(*
SPDX-FileCopyrightText: © 2026 Oleksandr Tiutyk <trofimich@gmail.com>
SPDX-License-Identifier: MIT
License: https://opensource.org/license/mit
*)

(*!
<summary>Writes run summaries and leaf failures to the ADS log.</summary>
<description>
Use in one task without reentry. The ADS backend has no established concurrent-call guarantee, even for
separate reporter instances. For multiple tasks use per-task in-memory reports or a synchronized backend.
Each callback submits at most one record. The ADS completion record includes counts and the first failed leaf name.
LastRunSummary includes the first failed leaf name and a bounded
version of its diagnostic. The summary and failed log writes are observable after the run. A failed
write does not change the test outcome. Individual ADS failure records are capped at 200 wide characters.
ReportRunStart clears all observations before attempting the start message.
</description>
*)

{attribute 'no_explicit_call' := 'do not call this function block directly'}
FUNCTION_BLOCK AdsLogReporter EXTENDS TOF_Core.Object IMPLEMENTS ITestReporter
VAR_STAT
	_ClassName : STRING := __POUNAME();
END_VAR
VAR
	_AdsLogger : TOF_Core.AdsLogger;
	_FirstFailureName : WSTRING;
	_FirstFailureDiagnostic : WSTRING(255);
	_LastRunSummary : TOF_Core.ERROR_MESSAGE;
	_FailedLogWriteCount : UDINT;
	_LastLogFailureMessage : TOF_Core.ERROR_MESSAGE;
END_VAR

(*!
<summary>Provides the implementation class name.</summary>
*)
{attribute 'monitoring' := 'call'}
PROPERTY ClassName : REFERENCE TO STRING
GET
ClassName REF= _ClassName;
END_GET
END_PROPERTY

(*!
<summary>Counts start, result and summary writes for which TryLogMessage returned FALSE.</summary>
<description>The count resets at ReportRunStart. A successful write does not confirm display in XAE.</description>
*)
{attribute 'monitoring' := 'call'}
PROPERTY FailedLogWriteCount : UDINT
GET
FailedLogWriteCount := _FailedLogWriteCount;
END_GET
END_PROPERTY

(*!
<summary>Borrows the last message whose ADS logger call returned FALSE.</summary>
<description>Empty until a write fails in the current run. Callers must not modify the returned storage.</description>
*)
{attribute 'monitoring' := 'call'}
PROPERTY LastLogFailureMessage : REFERENCE TO TOF_Core.ERROR_MESSAGE
GET
LastLogFailureMessage REF= _LastLogFailureMessage;
END_GET
END_PROPERTY

(*!
<summary>Borrows the summary created at ReportRunEnd regardless of its ADS write status.</summary>
<description>Empty after ReportRunStart until ReportRunEnd. Callers must not modify the returned storage.</description>
*)
{attribute 'monitoring' := 'call'}
PROPERTY LastRunSummary : REFERENCE TO TOF_Core.ERROR_MESSAGE
GET
LastRunSummary REF= _LastRunSummary;
END_GET
END_PROPERTY

(*!
<summary>Submits one ADS message and records a FALSE result from the logger.</summary>
<description>The count saturates at the largest UDINT. The copied text remains available until the next start.</description>
*)
METHOD PRIVATE logMessage
VAR_INPUT
	category : TOF_Core.LOG_CATEGORY;
END_VAR
VAR_IN_OUT CONSTANT
	message : TOF_Core.ERROR_MESSAGE;
END_VAR
IF TryWriteMessage(category := category, message := message) THEN
	RETURN;
END_IF

IF _FailedLogWriteCount < TOF_Core.UnsignedInt32.MAX_VALUE THEN
	_FailedLogWriteCount := _FailedLogWriteCount + 1;
END_IF

_LastLogFailureMessage := message;
END_METHOD

(*!
<summary>Provides the library namespace.</summary>
*)
{attribute 'monitoring' := 'call'}
PROPERTY NamespaceName : REFERENCE TO STRING
GET
NamespaceName REF= CurrentNamespace.Name;
END_GET
END_PROPERTY

(*!
<summary>Logs leaf counts and the first failed leaf name and retains its diagnostic for online inspection.</summary>
<description>The retained summary also includes a bounded first-failure diagnostic and survives a rejected ADS write.</description>
*)
METHOD ReportRunEnd
VAR_INPUT
	totalTests : TOF_Core.DINT_LENGTH;
	passedTests : TOF_Core.DINT_LENGTH;
	failedTests : TOF_Core.DINT_LENGTH;
	skippedTests : TOF_Core.DINT_LENGTH;
	duration : TIME;
END_VAR
VAR
	logSummary : WSTRING(255);
	logRecord : TOF_Core.ERROR_MESSAGE;
	summary : WSTRING(255);
END_VAR
summary := TOF_Core.WideStrings.Concat255(
	"[TOF_Testing] Finished: ", TO_WSTRING(passedTests), " passed, ",
	TO_WSTRING(failedTests), " failed, ", TO_WSTRING(skippedTests), " skipped"
);

logSummary := summary;

IF failedTests > 0 AND_THEN _FirstFailureDiagnostic <> "" THEN
	TOF_Core.WideStrings.AppendFit255(logSummary, " | First failed test: ", _FirstFailureName);
	TOF_Core.WideStrings.AppendFit255(summary, " | First failure: ", _FirstFailureDiagnostic);
END_IF

_LastRunSummary := summary;
logRecord := logSummary;
logMessage(category := TOF_Core.LOG_CATEGORY.INFORMATION, message := logRecord);
END_METHOD

(*!
<summary>Resets per-run observations and logs the number of configured leaf tests.</summary>
<description>A failed start-message write counts toward the new run.</description>
*)
METHOD ReportRunStart
VAR_INPUT
	testCount : TOF_Core.DINT_LENGTH;
END_VAR
VAR
	diagnostic : TOF_Core.ERROR_MESSAGE;
END_VAR
_FirstFailureName := "";
_FirstFailureDiagnostic := "";
_LastRunSummary := "";
_FailedLogWriteCount := 0;
_LastLogFailureMessage := "";

diagnostic := TOF_Core.WideStrings.Concat255(
	"[TOF_Testing] Starting ", TO_WSTRING(testCount), " tests"
);

logMessage(category := TOF_Core.LOG_CATEGORY.INFORMATION, message := diagnostic);
END_METHOD

(*!
<summary>Logs a failed leaf with its group path and caches the first failure for the summary.</summary>
<description>
The individual ADS record uses up to 200 wide characters to leave room below the native ADS text limit.
The retained summary includes the leaf name and the beginning of its diagnostic.
</description>
<param name="testName">Individual name bounded to 80 wide characters, matching INamed.</param>
*)
METHOD ReportTestCaseResult
VAR_INPUT
	groupPath : WSTRING(255);
	testName : WSTRING;
	outcome : TEST_OUTCOME;
	duration : TIME;
END_VAR
VAR_IN_OUT CONSTANT
	message : TOF_Core.ERROR_MESSAGE;
END_VAR
VAR
	shortDiagnostic : WSTRING(200);
	diagnostic : TOF_Core.ERROR_MESSAGE;
END_VAR
IF outcome <> TEST_OUTCOME.PASSED
	AND_THEN outcome <> TEST_OUTCOME.FAILED
	AND_THEN outcome <> TEST_OUTCOME.SKIPPED
THEN
	TOF_Core.Exceptions.ThrowArgumentValueNotSupported(
		sourceNamespaceName := NamespaceName,
		sourceClassName := ClassName,
		sourcePOUName := __POUNAME(),
		sourcePosition := __POSITION(),
		argumentName := 'outcome',
		argumentValue := outcome
	);
END_IF

IF outcome <> TEST_OUTCOME.FAILED THEN
	RETURN;
END_IF

IF _FirstFailureDiagnostic = "" THEN
	_FirstFailureName := testName;

	IF _FirstFailureName = "" THEN
		_FirstFailureName := "<unnamed>";
	END_IF

	_FirstFailureDiagnostic := TOF_Core.WideStrings.Concat255(_FirstFailureName, ": ");
	TOF_Core.WideStrings.AppendFit(targetString := _FirstFailureDiagnostic, sourceString := message);
END_IF

shortDiagnostic := "[TOF_Testing] ";

IF groupPath <> "" THEN
	TOF_Core.WideStrings.AppendFit255(shortDiagnostic, groupPath, "/");
END_IF

TOF_Core.WideStrings.AppendFit255(shortDiagnostic, testName, ": ");
TOF_Core.WideStrings.AppendFit(targetString := shortDiagnostic, sourceString := message);
diagnostic := shortDiagnostic;

logMessage(category := TOF_Core.LOG_CATEGORY.ERROR, message := diagnostic);
END_METHOD

(*!
<summary>Reports instance storage without separately allocated payloads.</summary>
*)
{attribute 'monitoring' := 'call'}
PROPERTY SelfSize : ULINT
GET
SelfSize := XSIZEOF(THIS^);
END_GET
END_PROPERTY

(*!
<summary>Submits one message to the ADS backend and reports whether the logger accepted it.</summary>
<description>
An override may replace the backend. It must return FALSE on rejection and must not raise an exception,
retry the write, or retain the borrowed message. TRUE does not confirm display in XAE.
</description>
*)
METHOD PROTECTED TryWriteMessage : BOOL
VAR_INPUT
	category : TOF_Core.LOG_CATEGORY;
END_VAR
VAR_IN_OUT CONSTANT
	message : TOF_Core.ERROR_MESSAGE;
END_VAR
TryWriteMessage := _AdsLogger.TryLogMessage(category := category, message := message);
END_METHOD

END_FUNCTION_BLOCK

(* stored: Version 1.1.0.1
   POU AdsLogReporter: Id {eb91e524-2438-48a4-9961-78fd9f56893c}, SpecialFunc None
   Property ClassName: Id {b69bfb0d-2ea3-4617-a4a6-eeca92a7fefb}
   Get Get: Id {b294ab84-b0af-46fc-8248-793022e91b31}
   Property FailedLogWriteCount: Id {159f9331-db53-4e73-ac02-b64bded2227f}
   Get Get: Id {c4093a24-5413-407f-ba52-31524df72870}
   Property LastLogFailureMessage: Id {96074640-3b0f-4b76-8958-405da4a01905}
   Get Get: Id {449ad356-f869-475c-b791-fe4802f56fac}
   Property LastRunSummary: Id {ac0e566d-a009-46ba-96e7-29baf150e0a0}
   Get Get: Id {3facb692-cf29-48f1-8262-90eea45ab450}
   Method logMessage: Id {c6cc75ab-d14a-43ed-82d8-6172cf95d6d4}
   Property NamespaceName: Id {307044c2-62a4-4bee-b8de-9823fa86f60c}
   Get Get: Id {92366a78-e137-465b-8ae9-cefa48f32002}
   Method ReportRunEnd: Id {f342d4f8-6bd1-4885-9c6d-263d40c86dfe}
   Method ReportRunStart: Id {e33e2cad-cdc4-4f26-9afe-7859394471ba}
   Method ReportTestCaseResult: Id {fef23984-ca74-4077-b47a-ac9e1f01e9b5}
   Property SelfSize: Id {0dd6e191-246a-483b-a793-65cba039133e}
   Get Get: Id {4b75b5da-6a57-48b6-ad20-c8ea20db62c7}
   Method TryWriteMessage: Id {7d405a37-57d8-443b-b1c8-999f47920d35} *)
